{region 'Documentation'}
(*!
<summary>Controlled I_Orchestrator boundary for Suite owner tests, without a scheduler.</summary>
<description>
Initialize records identity, collection bounds and child identities while the owner is still
initializing. Execute records task assignment and pre-child-call states. SetObservation supplies deliberate
responses between owner cycles; no child requests, reservations or state machine are copied.
The test supplies coherent child observations separately through the concrete Suite adapter.
</description>
*)
{endregion}
FUNCTION_BLOCK SuiteOrchestratorDouble IMPLEMENTS I_Orchestrator
VAR
    FAcceptInitialization : BOOL := TRUE;
    FInitialized : BOOL;
    FInitializeCount : UINT;
    FExecuteCount : UINT;
    FFirstChildStateAtExecute : E_State;
    FLastChildStateAtExecute : E_State;
    FCurrentTask : E_OrchestratorTask;
    FCollection : I_OrchestratableCollection;
    FName : STRING(GVL_Constants.NameLength);
    FResourceName : STRING(GVL_Constants.ResourceNameLength);
    FFirstIndex : DINT;
    FLastIndex : DINT;
    FChildCount : UINT;
    FFirstChild : I_Orchestratable;
    FLastChild : I_Orchestratable;
    FReady : BOOL;
    FResult : E_Result;
    FResetFinished : BOOL;
    FAbortFinished : BOOL;
    FExecutionFinished : BOOL;
END_VAR

{region 'Documentation'}
(*!
<summary>Clears observations before owner initialization and selects only the initialization outcome.</summary>
*)
{endregion}
METHOD PUBLIC BeginScenario
VAR_INPUT
    AcceptInitialization : BOOL := TRUE; //! Scripted acceptance returned by subsequent Initialize calls.
END_VAR
FAcceptInitialization := AcceptInitialization;
FInitialized := FALSE;
FInitializeCount := 0;
FExecuteCount := 0;
FFirstChildStateAtExecute := E_State.Uninitialized;
FLastChildStateAtExecute := E_State.Uninitialized;
FCurrentTask := E_OrchestratorTask.Idle;
FCollection := 0;
FName := '';
FResourceName := '';
FFirstIndex := 0;
FLastIndex := 0;
FChildCount := 0;
FFirstChild := 0;
FLastChild := 0;
SetObservation(Ready := FALSE);
END_METHOD

{region 'Documentation'}
(*!
<summary>Population observed synchronously inside Initialize.</summary>
*)
{endregion}
{attribute 'monitoring' := 'call'}
PROPERTY PUBLIC ChildCount : UINT //! Population observed synchronously inside Initialize.
GET
ChildCount := FChildCount;
END_GET
END_PROPERTY

{region 'Documentation'}
(*!
<summary>The exact collection interface supplied by the owner.</summary>
*)
{endregion}
{attribute 'monitoring' := 'variable'}
PROPERTY PUBLIC Collection : I_OrchestratableCollection //! The exact collection interface supplied by the owner.
GET
Collection := FCollection;
END_GET
END_PROPERTY

{region 'Documentation'}
(*!
<summary>Last task supplied by the owner.</summary>
*)
{endregion}
{attribute 'monitoring' := 'call'}
PROPERTY PUBLIC CurrentTask : E_OrchestratorTask //! Last task supplied by the owner.
GET
CurrentTask := FCurrentTask;
END_GET
END_PROPERTY

{region 'Documentation'}
(*!
<summary>Records the owner task and current child states; no observations are changed or child commands sent.</summary>
*)
{endregion}
METHOD PUBLIC Execute
VAR_INPUT
    Task : E_OrchestratorTask; //! Owner-assigned task to record; this double does not execute or request children.
END_VAR
FCurrentTask := Task;
FExecuteCount := FExecuteCount + 1;
IF FFirstChild <> 0 THEN
    FFirstChildStateAtExecute := FFirstChild.State;
END_IF;
IF FLastChild <> 0 THEN
    FLastChildStateAtExecute := FLastChild.State;
END_IF;
END_METHOD

{region 'Documentation'}
(*!
<summary>Number of cyclic helper calls.</summary>
*)
{endregion}
{attribute 'monitoring' := 'call'}
PROPERTY PUBLIC ExecuteCount : UINT //! Number of cyclic helper calls.
GET
ExecuteCount := FExecuteCount;
END_GET
END_PROPERTY

{region 'Documentation'}
(*!
<summary>First occupied interface observed inside Initialize.</summary>
*)
{endregion}
{attribute 'monitoring' := 'variable'}
PROPERTY PUBLIC FirstChild : I_Orchestratable //! First occupied interface observed inside Initialize.
GET
FirstChild := FFirstChild;
END_GET
END_PROPERTY

{region 'Documentation'}
(*!
<summary>First child state observed by the helper before concrete child calls.</summary>
*)
{endregion}
{attribute 'monitoring' := 'call'}
PROPERTY PUBLIC FirstChildStateAtExecute : E_State //! First child state observed by the helper before concrete child calls.
GET
FirstChildStateAtExecute := FFirstChildStateAtExecute;
END_GET
END_PROPERTY

{region 'Documentation'}
(*!
<summary>Lower bound observed synchronously inside Initialize.</summary>
*)
{endregion}
{attribute 'monitoring' := 'call'}
PROPERTY PUBLIC FirstIndex : DINT //! Lower bound observed synchronously inside Initialize.
GET
FirstIndex := FFirstIndex;
END_GET
END_PROPERTY

{region 'Documentation'}
(*!
<summary>Records and immediately queries the collection handed over by the owner; never executes children.</summary>
*)
{endregion}
METHOD PUBLIC Initialize : BOOL //! Scripted initialization acceptance; the supplied collection is queried regardless of that response.
VAR_INPUT
    Collection : I_OrchestratableCollection; //! Nonzero borrowed collection queried immediately and retained; keep the collection and children alive.
    Name : STRING(GVL_Constants.NameLength); //! Owner diagnostic name retained by the double.
    ResourceName : STRING(GVL_Constants.ResourceNameLength) := ''; //! Owner diagnostic resource retained by the double.
END_VAR
FInitializeCount := FInitializeCount + 1;
FCollection := Collection;
FName := Name;
FResourceName := ResourceName;
FFirstIndex := Collection.ChildArrayLowerBound;
FLastIndex := Collection.ChildArrayUpperBound;
FChildCount := Collection.ChildCount;
IF FChildCount > 0 THEN
    FFirstChild := Collection.GetChild(Index := FFirstIndex);
    FLastChild := Collection.GetChild(Index := FFirstIndex + UINT_TO_DINT(FChildCount) - 1);
END_IF;
FInitialized := FAcceptInitialization;
Initialize := FInitialized;
END_METHOD

{region 'Documentation'}
(*!
<summary>Number of owner initialization calls.</summary>
*)
{endregion}
{attribute 'monitoring' := 'call'}
PROPERTY PUBLIC InitializeCount : UINT //! Number of owner initialization calls.
GET
InitializeCount := FInitializeCount;
END_GET
END_PROPERTY

{region 'Documentation'}
(*!
<summary>Scripted Abort completion.</summary>
*)
{endregion}
{attribute 'monitoring' := 'call'}
PROPERTY PUBLIC IsAbortFinished : BOOL //! Scripted Abort completion.
GET
IsAbortFinished := FAbortFinished;
END_GET
END_PROPERTY

{region 'Documentation'}
(*!
<summary>Scripted execution completion.</summary>
*)
{endregion}
{attribute 'monitoring' := 'call'}
PROPERTY PUBLIC IsExecutionFinished : BOOL //! Scripted execution completion.
GET
IsExecutionFinished := FExecutionFinished;
END_GET
END_PROPERTY

{region 'Documentation'}
(*!
<summary>Accepted initialization response.</summary>
*)
{endregion}
{attribute 'monitoring' := 'call'}
PROPERTY PUBLIC IsInitialized : BOOL //! Accepted initialization response.
GET
IsInitialized := FInitialized;
END_GET
END_PROPERTY

{region 'Documentation'}
(*!
<summary>Scripted child readiness summary.</summary>
*)
{endregion}
{attribute 'monitoring' := 'call'}
PROPERTY PUBLIC IsReady : BOOL //! Scripted child readiness summary.
GET
IsReady := FReady;
END_GET
END_PROPERTY

{region 'Documentation'}
(*!
<summary>Whether the owner currently assigns Reset.</summary>
*)
{endregion}
{attribute 'monitoring' := 'call'}
PROPERTY PUBLIC IsResetActive : BOOL //! Whether the owner currently assigns Reset.
GET
IsResetActive := FCurrentTask = E_OrchestratorTask.Reset;
END_GET
END_PROPERTY

{region 'Documentation'}
(*!
<summary>Scripted Reset completion.</summary>
*)
{endregion}
{attribute 'monitoring' := 'call'}
PROPERTY PUBLIC IsResetFinished : BOOL //! Scripted Reset completion.
GET
IsResetFinished := FResetFinished;
END_GET
END_PROPERTY

{region 'Documentation'}
(*!
<summary>Last occupied interface observed inside Initialize.</summary>
*)
{endregion}
{attribute 'monitoring' := 'variable'}
PROPERTY PUBLIC LastChild : I_Orchestratable //! Last occupied interface observed inside Initialize.
GET
LastChild := FLastChild;
END_GET
END_PROPERTY

{region 'Documentation'}
(*!
<summary>Last child state observed by the helper before concrete child calls.</summary>
*)
{endregion}
{attribute 'monitoring' := 'call'}
PROPERTY PUBLIC LastChildStateAtExecute : E_State //! Last child state observed by the helper before concrete child calls.
GET
LastChildStateAtExecute := FLastChildStateAtExecute;
END_GET
END_PROPERTY

{region 'Documentation'}
(*!
<summary>Capacity upper bound observed synchronously inside Initialize.</summary>
*)
{endregion}
{attribute 'monitoring' := 'call'}
PROPERTY PUBLIC LastIndex : DINT //! Capacity upper bound observed synchronously inside Initialize.
GET
LastIndex := FLastIndex;
END_GET
END_PROPERTY

{region 'Documentation'}
(*!
<summary>Diagnostic identity supplied by the owner.</summary>
*)
{endregion}
{attribute 'monitoring' := 'variable'}
PROPERTY PUBLIC OwnerName : STRING(GVL_Constants.NameLength) //! Diagnostic identity supplied by the owner.
GET
OwnerName := FName;
END_GET
END_PROPERTY

{region 'Documentation'}
(*!
<summary>Diagnostic resource supplied by the owner.</summary>
*)
{endregion}
{attribute 'monitoring' := 'variable'}
PROPERTY PUBLIC ResourceName : STRING(GVL_Constants.ResourceNameLength) //! Diagnostic resource supplied by the owner.
GET
ResourceName := FResourceName;
END_GET
END_PROPERTY

{region 'Documentation'}
(*!
<summary>Scripted helper technical result.</summary>
*)
{endregion}
{attribute 'monitoring' := 'call'}
PROPERTY PUBLIC Result : E_Result //! Scripted helper technical result.
GET
Result := FResult;
END_GET
END_PROPERTY

{region 'Documentation'}
(*!
<summary>Supplies the interface response for the next owner call; defaults describe unfinished neutral work.</summary>
*)
{endregion}
METHOD PUBLIC SetObservation
VAR_INPUT
    Ready : BOOL; //! Scripted readiness returned to the owner.
    Result : E_Result := E_Result.NotEvaluated; //! Scripted helper technical result returned to the owner.
    ResetFinished : BOOL := FALSE; //! Scripted Reset-completion signal returned to the owner.
    AbortFinished : BOOL := FALSE; //! Scripted Abort-completion signal returned to the owner.
    ExecutionFinished : BOOL := FALSE; //! Scripted execution-completion signal returned to the owner.
END_VAR
FReady := Ready;
FResult := Result;
FResetFinished := ResetFinished;
FAbortFinished := AbortFinished;
FExecutionFinished := ExecutionFinished;
END_METHOD

END_FUNCTION_BLOCK

(* stored: Version 1.1.0.1
   POU SuiteOrchestratorDouble: Id {55b7b544-5c0e-41b4-9a1c-3c3d7a542c1a}, SpecialFunc None
   Folder Internal: Id {4c1a09d9-e984-4d97-a5a1-3f6de02e8ccf}
   Method BeginScenario: Id {aef1639a-7b7c-4fe7-81cb-1f222d311e18}
   Property ChildCount: Id {bae0f3d4-9656-453d-ae93-7c4b0f855be1}
   Get Get: Id {3a0f0ff9-0622-4076-9895-54586d44fc0a}
   Property Collection: Id {5938fd68-0b28-41f2-96fe-cd3b1f3fcce7}
   Get Get: Id {269283e5-a782-4a06-a420-2672cf24ec3d}
   Property CurrentTask: Id {bdaac40f-a4bc-4c17-a1f6-17bb128dcb7e}
   Get Get: Id {5f5ab9b6-1685-4717-8710-700b2879cc0b}
   Method Execute: Id {57263bee-e8bf-4efc-b2af-97e29b65daf1}
   Property ExecuteCount: Id {4a647fd0-3c53-4b05-acf2-fe263aabd681}
   Get Get: Id {65e0475d-70ad-471b-bf36-f46ab855ffde}
   Property FirstChild: Id {10eed8a1-b409-4362-8a15-8deb57cf5c41}
   Get Get: Id {97030e9e-872c-4b94-be8c-b2474f7f4e73}
   Property FirstChildStateAtExecute: Id {053a285a-f919-468d-8fbe-5b8dbbeba05e}
   Get Get: Id {eeb2ba4e-cf95-44bc-ab58-813f3ec6e8ca}
   Property FirstIndex: Id {c1e2a98e-eabe-4f9a-b5b4-69b12cf27f83}
   Get Get: Id {f923fced-27d9-407a-88d9-d3169ae2cbf0}
   Method Initialize: Id {ae1adbac-4d4b-4a86-b04b-5528b94496f3}
   Property InitializeCount: Id {ef016cc3-4acb-48ae-bffa-bb8adef5af2e}
   Get Get: Id {a3539587-b914-47ce-8ee2-7952f2e54c7e}
   Property IsAbortFinished: Id {ee43daa6-a119-4efd-b566-37639efa8cb1}
   Get Get: Id {00df052e-ac4d-4ec7-801d-30a17a1cc35e}
   Property IsExecutionFinished: Id {08f024a8-72cc-44cb-820c-0f31eb90c78d}
   Get Get: Id {6f41bb1a-7103-4e4a-94e9-b5cf96db0f44}
   Property IsInitialized: Id {e4e44681-9a95-4413-9632-b29097800a72}
   Get Get: Id {533dc622-b16d-459c-8a77-d24fb18ba428}
   Property IsReady: Id {410035f4-35b7-4872-971e-0ab11afe44f1}
   Get Get: Id {4506be1d-2502-4272-8754-b16eb40bac6b}
   Property IsResetActive: Id {575a31fb-8132-4477-baaa-32ea5e345c21}
   Get Get: Id {72249477-7852-48a3-b54c-4cdfa68d0bb5}
   Property IsResetFinished: Id {4f3900db-248c-4bfa-9e37-204b1daa14ef}
   Get Get: Id {5f5ea8be-8e04-4526-b28e-89139384bcb5}
   Property LastChild: Id {eaae123c-7d81-48b6-a43e-b91f2ee42a70}
   Get Get: Id {389ee9ad-5640-4a55-b293-972d1d481d19}
   Property LastChildStateAtExecute: Id {e95a4bb1-40a5-4a92-a794-5ba274b874fe}
   Get Get: Id {690d19e1-1f52-458c-af71-06e7a50b5600}
   Property LastIndex: Id {c0d9dc8c-bee4-442f-9274-20fcf4e514f9}
   Get Get: Id {ecd4d208-7fcd-4675-bea1-b497e0bf6e08}
   Property OwnerName: Id {9b64f83f-d2d7-4d0d-b919-37b9c386afb2}
   Get Get: Id {6d514031-6ff3-4551-ac81-a0f8814b53db}
   Property ResourceName: Id {93e22e8c-f12f-47e5-b983-38cd268d3f42}
   Get Get: Id {b0494098-abce-4a00-bf34-25a479644c0f}
   Property Result: Id {60d84426-0fe8-47cd-a448-f7e2db82dae1}
   Get Get: Id {5247e920-ebd3-4598-bcda-19d0257cdaf6}
   Method SetObservation: Id {63041564-ffdf-4eb0-ae93-a472c89d4a4a} *)
